TYPE "UDT_Service_ProcedureRawDataMedium"
VERSION : 0.1
   STRUCT
      procedure : Array[0..15] of "UDT_MTP_ProcedureExtended";
   END_STRUCT;

END_TYPE

